(* IEC 61131-3 sources: STAR-PLC-Agent/results/raw/codex_matrix_resume_20261114/codex_terra/PUB013/formal/attempt_0001, 1 file *)

(* ---- candidate.st ---- *)
FUNCTION_BLOCK FB_Task
VAR_INPUT
    OCCUPANCY_DETECTED : BOOL;
    ENERGY_SAVING_MODE : BOOL;
    HVAC_MODE_SELECTOR : INT;
END_VAR
VAR_OUTPUT
    SUPPLY_FAN_RUN : BOOL := FALSE;
    TEMP_SETPOINT_ADJUST : INT := 0;
END_VAR
VAR
    FanDelay : TON;
END_VAR

FanDelay(IN := OCCUPANCY_DETECTED AND (HVAC_MODE_SELECTOR <> 3), PT := T#30s);
SUPPLY_FAN_RUN := FanDelay.Q;

CASE HVAC_MODE_SELECTOR OF
    0:
        IF OCCUPANCY_DETECTED THEN
            TEMP_SETPOINT_ADJUST := 0;
        ELSIF ENERGY_SAVING_MODE THEN
            TEMP_SETPOINT_ADJUST := 3;
        ELSE
            TEMP_SETPOINT_ADJUST := 2;
        END_IF;
    1:
        IF OCCUPANCY_DETECTED THEN
            TEMP_SETPOINT_ADJUST := 0;
        ELSE
            TEMP_SETPOINT_ADJUST := 1;
        END_IF;
    2:
        IF OCCUPANCY_DETECTED THEN
            TEMP_SETPOINT_ADJUST := 0;
        ELSE
            TEMP_SETPOINT_ADJUST := 4;
        END_IF;
    3:
        TEMP_SETPOINT_ADJUST := 4;
ELSE
    TEMP_SETPOINT_ADJUST := 0;
END_CASE;
END_FUNCTION_BLOCK
